FUNCTION_BLOCK FB_LogRecordExporter_HTTP EXTENDS FB_LogRecordExporter_Base
VAR_OUTPUT
	currentState: E_HttpExporterState;
	statusCode: UINT;  // the HTTP status code received for the last completed request
END_VAR

VAR
	_execute: BOOL;
	_urlParsed: BOOL;
	_endpoint: ST_HttpEndpoint;
	_len: UDINT;
	_execRTrig: R_TRIG;
	_pString: POINTER TO STRING;
	_jsonVal: SJsonValue;
	_computedState: E_HttpExporterState;
	_failureReason: E_LogRecordExporterFailureReason;
	_serializationFailureReason: E_ProtoJsonSerializerFailureReason;
	_serializer: FB_LogRecordProtoJsonSerializer;
	_client: FB_IotHttpClient;
	_request: FB_IotHttpRequest;
	_header: FB_IotHttpHeaderFieldMap;
END_VAR

THIS^.tick(failureReason=>THIS^._callFailureReason);

METHOD export: BOOL
VAR_IN_OUT
	logRecords: FB_LogRecordQueue;
END_VAR
VAR_INPUT
	count: UDINT;
END_VAR
VAR_OUTPUT
	failureReason: E_LogRecordExporterFailureReason;
END_VAR
// Prepare a completed exporter to accept the next batch immediately.
IF THIS^.currentState = E_HttpExporterState.done OR THIS^.currentState = E_HttpExporterState.error THEN
	THIS^.currentState := E_HttpExporterState.idle;
	THIS^._computedState := E_HttpExporterState.idle;
END_IF
export := SUPER^.export(
	logRecords:=logRecords,
	count:=count,
	failureReason=>failureReason
);
IF export THEN
	THIS^._failureReason := E_LogRecordExporterFailureReason.NA;
	THIS^._serializationFailureReason := E_ProtoJsonSerializerFailureReason.NA;
END_IF
END_METHOD

(*
	Releases a payload buffer that is still in flight. The FB_IotHttpRequest reading it is
	destroyed with this instance, so nothing uses the buffer afterwards. TwinCAT then
	runs FB_LogRecordExporter_Base.FB_Exit, which releases the queued records.
*)
METHOD FB_Exit : BOOL
VAR_INPUT
	bInCopyCode: BOOL;  // TRUE: the instance is being copied during an online change
END_VAR
// during an online change the copy keeps the buffer, so it must not be released here
IF NOT bInCopyCode AND _pString <> 0 THEN
	__DELETE(_pString);
	_pString := 0;
END_IF
END_METHOD

//FB_Init is always available implicitly and it is used primarily for initialization.
//The return value is not evaluated. For a specific influence, you can also declare the
//methods explicitly and provide additional code there with the standard initialization
//code. You can evaluate the return value.
METHOD FB_Init: BOOL
VAR_INPUT
	bInitRetains: BOOL; // TRUE: the retain variables are initialized (reset warm / reset cold)
	bInCopyCode: BOOL;  // TRUE: the instance will be copied to the copy code afterward (online change)
	url: T_MaxString;  // full endpoint URL, e.g. 'http://192.168.1.10:4318/v1/logs'
	bNoServerCertCheck: BOOL := FALSE;  // allow HTTPS connections to servers with self-signed certificates
END_VAR
THIS^.currentState := E_HttpExporterState.idle;
THIS^._computedState := E_HttpExporterState.idle;

THIS^._urlParsed := F_ParseHttpUrl(url:=url, endpoint=>THIS^._endpoint);

THIS^._client.sHostName := THIS^._endpoint.host;
THIS^._client.nHostPort := THIS^._endpoint.port;
THIS^._client.bKeepAlive := TRUE;
THIS^._client.tConnectionTimeout := T#10S;
IF THIS^._endpoint.useTls THEN
	THIS^._client.stTLS.bNoServerCertCheck := bNoServerCertCheck;
END_IF

THIS^._request.sContentType := 'application/json';
END_METHOD

METHOD isBusy : BOOL
isBusy := THIS^._exportActive;
END_METHOD

METHOD tick : BOOL
VAR_OUTPUT
	failureReason: E_LogRecordExporterFailureReason;
END_VAR
tick := TRUE;
failureReason := E_LogRecordExporterFailureReason.NA;

_execute := THIS^._exportActive;
_execRTrig(CLK := _execute AND_THEN THIS^._records.count > 0);

CASE currentState OF
	E_HttpExporterState.idle:
		IF _execRTrig.Q THEN
			_failureReason := E_LogRecordExporterFailureReason.NA;
			_serializationFailureReason := E_ProtoJsonSerializerFailureReason.NA;
			IF NOT THIS^._urlParsed THEN
				_failureReason := E_LogRecordExporterFailureReason.HTTP_URL_PARSE_FAILURE;
				_computedState := E_HttpExporterState.error;
			ELSE
				_computedState := E_HttpExporterState.serializing;
			END_IF
		END_IF

	E_HttpExporterState.serializing:
		// Serialize the batch and buffer the LogsData document as a byte array payload.
		IF NOT _serializer.serializeLogsData(
			logRecords:=THIS^._records,
			failureReason=>_serializationFailureReason
		) THEN
			_failureReason := E_LogRecordExporterFailureReason.SERIALIZATION_FAILURE;
			_computedState := E_HttpExporterState.error;
		ELSE
			_jsonVal := _serializer.jsonValue;
			IF _jsonVal = 0 OR_ELSE NOT _serializer.parser.IsObject(_jsonVal) THEN
				_failureReason := E_LogRecordExporterFailureReason.SERIALIZATION_FAILURE;
				_computedState := E_HttpExporterState.error;
			ELSE
				_len := _serializer.parser.GetJsonLength(_jsonVal);  // includes the null terminating character
				IF _len = 0 THEN
					_failureReason := E_LogRecordExporterFailureReason.SERIALIZATION_FAILURE;
					_computedState := E_HttpExporterState.error;
				ELSE
					_pString := __NEW(BYTE, _len);
					IF _pString = 0 THEN
						_failureReason := E_LogRecordExporterFailureReason.BUFFER_ALLOCATION_FAILURE;
						_computedState := E_HttpExporterState.error;
					ELSE
						_serializer.parser.CopyJson(_jsonVal, _pString^, _len);
						_computedState := E_HttpExporterState.sending;
					END_IF
				END_IF
			END_IF
		END_IF

	E_HttpExporterState.sending:
		IF NOT _request.bBusy THEN
			IF _request.SendRequest(
				sUri := THIS^._endpoint.path,
				fbClient := THIS^._client,
				eRequestType := ETcIotHttpRequestType.HTTP_POST,
				pContent := _pString,
				nContentSize := _len - 1,
				fbHeader := THIS^._header
			) THEN
				_computedState := E_HttpExporterState.waiting;
			ELSE
				IF _pString <> 0 THEN __DELETE(_pString); _pString := 0; END_IF
				_failureReason := E_LogRecordExporterFailureReason.HTTP_REQUEST_FAILURE;
				_computedState := E_HttpExporterState.error;
			END_IF
		END_IF

	E_HttpExporterState.waiting:
		IF NOT _request.bBusy THEN
			_computedState := E_HttpExporterState.processing;
		END_IF

	E_HttpExporterState.processing:
		IF _request.bError THEN
			IF _pString <> 0 THEN __DELETE(_pString); _pString := 0; END_IF
			_failureReason := E_LogRecordExporterFailureReason.HTTP_REQUEST_FAILURE;
			_computedState := E_HttpExporterState.error;
		ELSE
			statusCode := _request.nStatusCode;
			IF statusCode < 200 OR_ELSE statusCode >= 300 THEN
				IF _pString <> 0 THEN __DELETE(_pString); _pString := 0; END_IF
				_failureReason := E_LogRecordExporterFailureReason.HTTP_STATUS_FAILURE;
				_computedState := E_HttpExporterState.error;
			ELSE
				IF _pString <> 0 THEN __DELETE(_pString); _pString := 0; END_IF
				_computedState := E_HttpExporterState.done;
			END_IF
		END_IF

	E_HttpExporterState.done:
		IF NOT _execute THEN
			_computedState := E_HttpExporterState.idle;
		END_IF
		THIS^.free();

	E_HttpExporterState.error:
		// Retain the failure until export accepts a new batch.
END_CASE

currentState := _computedState;

IF currentState = E_HttpExporterState.done
	OR_ELSE currentState = E_HttpExporterState.error THEN
	THIS^.free();
END_IF

THIS^._client.Execute();

IF currentState = E_HttpExporterState.error THEN
	tick := FALSE;
	failureReason := _failureReason;
END_IF
END_METHOD

END_FUNCTION_BLOCK

(* stored: Version 1.1.0.1
   POU FB_LogRecordExporter_HTTP: Id {94541c0f-c88a-4178-bb34-d3823fe70965}, SpecialFunc None
   Method export: Id {c1e9c3db-bbd6-4dba-b7b4-d5219023c6d6}
   Method FB_Exit: Id {5bddf7d2-c571-4f61-a937-216ec416b501}
   Method FB_Init: Id {62b2e312-9bed-4019-8a5b-4e0d487d8a0a}
   Method isBusy: Id {40cc32d7-f759-46ec-80dd-15e4415f71f5}
   Method tick: Id {9b2355dd-f7b1-4921-8536-533aebcd5760} *)
